(* IEC 61131-3 sources: POMIRTS_lab3/AS/Library/brsystem, 2 files *)

(* ---- brsystem.fun ---- *)
(********************************************************************
 * COPYRIGHT -- Bernecker + Rainer
 ********************************************************************
 * Library: brsystem
 * File: brsystem.fun
 * Author: B+R
 ********************************************************************
 * Functions and function blocks of library brsystem
 ********************************************************************)

FUNCTION_BLOCK MEMInfo				(*returns information about the memory areas available on the system*)
	VAR_INPUT
		enable	:BOOL;				(*enables execution*)
	END_VAR
	VAR_OUTPUT
		status	:UINT;				(*execution status: ERR_OK, ERR_FUB_ENABLE_FALSE, 0xXXXX = see help*)
		FreeUSR_Ram	:UDINT;			(*SG3: free memory in USER RAM SG4: free memory in SRAM (Userram)*)
		FreeSYSTEM	:UDINT;			(*SG3: free system memory SG4: not used, always 0*)
		FreeUSR_Prom	:UDINT;		(*SG3: free memory in USER PROM SG4: free memory of HD where RPSHD is located*)
		FreeSYS_Prom	:UDINT;		(*SG3: free memory in system PROM SG4: free memory of HD where RPSHD is located*)
		FreeFIX_Ram	:UDINT;			(*SG3: free memory in FIX RAM SG4: not used, always 0*)
		FreeTMP_Ram	:UDINT;			(*SG3: free temporary memory in RAM SG4: free memory in DRAM*)
		FreeMEMCARD	:UDINT;			(*SG3: free memory on MEMCARD SG4: not used, always 0*)
	END_VAR
END_FUNCTION_BLOCK

FUNCTION_BLOCK MEMxInfo				(*returns information about the memory areas available in the system; asynchronous execution*)
	VAR_INPUT
		enable	:BOOL;   			(*enables execution*)
		mem_typ	:UDINT;				(*memory type: brDRAM, brUSRRAM, brSYSROM, brUSRROM*)
	END_VAR
	VAR_OUTPUT
		status	:UINT;				(*execution status: ERR_OK, ERR_FUB_ENABLE_FALSE, ERR_FUB_BUSY, 0xXXXX = see help*)
		MemSize	:UDINT;				(*total memory size in bytes*)
		FreeMemSize	:UDINT;			(*size of available memory in bytes*)
		BiggestFreeBlockSize	:UDINT;	(*size of the largest available block in memory in bytes*)
	END_VAR
	VAR
		i_state	:UINT;				(*internal variable*)
		i_result	:UINT;			(*internal variable*)
		i_tmp	:UDINT;				(*internal variable*)
	END_VAR
END_FUNCTION_BLOCK

FUNCTION_BLOCK SysInfo				(*returns information about the target system*)
	VAR_INPUT
		enable	:BOOL;				(*enables execution*)
	END_VAR
	VAR_OUTPUT
		init_reason	:USINT;			(*reason for initialization*)
		init_count	:USINT;			(*SG3: the value is increased by every INIT (warm restart) SG4: not used, always 0*)
		tick_count	:UDINT;			(*tick count*)
		version	:UDINT;				(*operating system version of the target system*)
	END_VAR
END_FUNCTION_BLOCK

FUNCTION_BLOCK RTInfo				(*returns runtime information about the software object*)
	VAR_INPUT
		enable	:BOOL;				(*enables execution*)
	END_VAR
	VAR_OUTPUT
		status	:UINT;				(*execution status: ERR_OK, ERR_FUB_ENABLE_FALSE, 0xXXXX = see help*)
		cycle_time	:UDINT;			(*cycle time in microsec*)
		init_reason	:SINT;			(*reason for initialization*)
		task_class	:SINT;			(*task class (SG3: #1 - #4 SG4: #1 - #8)*)
	END_VAR
END_FUNCTION_BLOCK

FUNCTION_BLOCK TARGETInfo			(*returns information about the target system used*)
	VAR_INPUT
		enable	:BOOL;				(*enables execution*)
		pOSVersion	:UDINT;			(*string given as a pointer (min. 7 char), where the os version is written*)
	END_VAR
	VAR_OUTPUT
		status	:UINT;				(*execution status: ERR_OK, ERR_FUB_ENABLE_FALSE, 0xXXXX = see help*)
		DataFormat	:USINT;			(*wether "big endian" or "little endian" ("TARGET_BIG_ENDIAN"/"TARGET_LITTLE_ENDIAN")*)
	END_VAR
END_FUNCTION_BLOCK

FUNCTION_BLOCK HWInfo				(*returns information about the hardware configuration*)
	VAR_INPUT
		enable	:BOOL;				(*enables execution*)
		first	:BOOL;				(*determines the hardware module on which the FUB is used 0/1 next/first*)
		pName	:UDINT;				(*string given as a pointer, where the name of the module is written*)
	END_VAR
	VAR_OUTPUT
		status	:UINT;				(*execution status: ERR_OK, ERR_FUB_ENABLE_FALSE, 0xXXXX = see help*)
		family	:USINT;				(*family designation*)
		usetype	:USINT;				(*hardware type*)
		module_typ	:UDINT;			(*module type*)
		master_no	:USINT;			(*logical number of the IO master, RIO master, CAN bus with CANIO*)
		slave_no	:USINT;			(*slave number*)
		module_adr	:USINT;			(*hardware module address (decimal)*)
		slot_no	:USINT;				(*slot of the first submodule found (decimal)*)
	END_VAR
	VAR
		next_vw_p	:UDINT;			(*internal variable*)
		last_modul_p	:UDINT;		(*internal variable*)
		next_entry_p	:UDINT;		(*internal variable*)
		next_entry_ix	:USINT;		(*internal variable*)
		next_slot_ix	:USINT;		(*internal variable*)
		last_rio_master	:USINT;		(*internal variable*)
	END_VAR
END_FUNCTION_BLOCK

FUNCTION_BLOCK SysconfInfo			(*returns the parameters for a sysconf entry*)
	VAR_INPUT
		enable	:BOOL;				(*enables execution*)
		pEntry	:UDINT;				(*string given as a pointer, where the name of the entry is written*)
		pValue	:UDINT;				(*string given as a pointer, where the value of the entry is copied*)
		value_len	:UDINT;			(*length of the "value-string"*)
	END_VAR
	VAR_OUTPUT
		status	:UINT;				(*execution status: ERR_OK, ERR_FUB_ENABLE_FALSE, 0xXXXX = see help*)
	END_VAR
END_FUNCTION_BLOCK

FUNCTION_BLOCK SysconfSet			(*sets the parameters for a sysconf entry*)
	VAR_INPUT
		enable	:BOOL;				(*enables execution*)
		pEntry	:UDINT;				(*string given as a pointer, where the name of the entry is written*)
		pNewValue	:UDINT;			(*string given as a pointer, where the new value of the entry is written*)
		option	:USINT;				(*sets the parameter volatile/permanent ("brSYSCONF_SET_VOLATILE"/"brSYSCONF_SET_NON_VOLATILE")*)
	END_VAR
	VAR_OUTPUT
		status	:UINT;				(*execution status: ERR_OK, ERR_FUB_ENABLE_FALSE, 0xXXXX = see help*)
	END_VAR
END_FUNCTION_BLOCK

FUNCTION_BLOCK BatteryInfo			(*returns the state of the battery*)
	VAR_INPUT
		enable	:BOOL;				(*enables execution*)
		pDevice	:UDINT;				(*device name given as a pointer*)
	END_VAR
	VAR_OUTPUT
		status	:UINT;				(*execution status: ERR_OK, ERR_FUB_ENABLE_FALSE, 0xXXXX = see help*)
		state	:USINT;				(*state of the battery*)
	END_VAR
END_FUNCTION_BLOCK

FUNCTION_BLOCK EXCInfo				(*returns information about the software object that triggered the exception*)
	VAR_INPUT
		enable	:BOOL;				(*enables execution*)
	END_VAR
	VAR_OUTPUT
		status	:UINT;				(*execution status: ERR_OK, ERR_FUB_ENABLE_FALSE, 0xXXXX = see help*)
		task_class	:UDINT;			(*task class in which the exception was triggered*)
		task_ident	:UDINT;			(*ID number of the software object that triggered the exception*)
	END_VAR
END_FUNCTION_BLOCK

FUNCTION_BLOCK ZYKVLenable			(*enables/disables the cycle time monitoring of software objects*)
	VAR_INPUT
		enable	:BOOL;				(*enables execution*)
		mode	:BOOL;				(*0/1 monitoring off/on*)
	END_VAR
	VAR_OUTPUT
		status	:UINT;				(*execution status: ERR_OK, ERR_FUB_ENABLE_FALSE, 0xXXXX = see help*)
	END_VAR
END_FUNCTION_BLOCK

FUNCTION_BLOCK PMemGet				(*reads data of len byte from the permanent memeory area beginning at offset*)
	VAR_INPUT
		enable	:BOOL;				(*enables execution*)
		offset	:UDINT;				(*offset within the permanent memory area*)
		len	 :UDINT;				(*length of data area to be read*)
		adress	:UDINT;				(*address where the read data is copied*)
	END_VAR
	VAR_OUTPUT
		status	:UINT;				(*execution status: ERR_OK, ERR_FUB_ENABLE_FALSE, 0xXXXX = see help*)
	END_VAR
END_FUNCTION_BLOCK

FUNCTION_BLOCK PMemPut				(*writes len bytes to the permanent memory area beginning at offset*)
	VAR_INPUT
		enable	:BOOL;				(*enables execution*)
		offset	:UDINT;				(*offset within the permanent memory area*)
		len	 :UDINT;				(*length of data area to be written*)
		adress	:UDINT;				(*address of the data to be written to the permanent memory area*)
	END_VAR
	VAR_OUTPUT
		status	:UINT;				(*execution status: ERR_OK, ERR_FUB_ENABLE_FALSE, 0xXXXX = see help*)
	END_VAR
END_FUNCTION_BLOCK

FUNCTION_BLOCK PMemSize				(*determines the size of permanent memory area in its existing configuration*)
	VAR_INPUT
		enable	:BOOL;				(*enables execution*)
	END_VAR
	VAR_OUTPUT
		status	:UINT;				(*execution status: ERR_OK, ERR_FUB_ENABLE_FALSE, 0xXXXX = see help*)
		size	:UDINT;				(*size of permanent memory area*)
	END_VAR
END_FUNCTION_BLOCK

(* ---- brsystem.var ---- *)
(********************************************************************
 * COPYRIGHT -- Bernecker + Rainer
 ********************************************************************
 * Library: brsystem
 * File: brsystem.var
 * Author: B+R
 ********************************************************************
 * Local variables of library brsystem
 ********************************************************************)

VAR CONSTANT
	brSYSCONF_SET_NON_VOLATILE	: BOOL	:= TRUE;	(*set permanent value*)
	brERR_INVALID_PARAMETER	: UINT	:= 27251;		(*invalid parameter transferred*)
	brSYSCONF_SET_VOLATILE	: BOOL	:= FALSE;		(*set non-permanent value*)
	INIT_REASON_WARMSTART	: SINT	:= 1;			(*warm restart boot information*)
	INIT_REASON_COLDSTART	: SINT	:= 2;			(*cold restart boot information*)
	brERR_INVALID_DEVICE	: UINT	:= 27250;		(*battery monitoring*)
	brAUTOMATION_RUNTIME	: USINT	:= 4;			(*series recognition*)
	TARGET_LITTLE_ENDIAN	: USINT	:= 1;			(*formatSpec*)
	INIT_REASON_DOWNLOAD	: SINT	:= 3;			(*download boot information*)
	INIT_REASON_UNKNOWN	: SINT	:= -1;				(*unknown boot information*)
	brBATTERY_MISSING	: USINT	:= 3;				(*battery monitoring*)
	TARGET_BIG_ENDIAN	: USINT	:= 2;				(*formatSpec*)
	brBATTERY_NOTEST	: USINT	:= 2;				(*battery monitoring*)
	brSYSTEM_MODULE	: USINT	:= 2;					(*usage recognition*)
	brPLUGIN_MODULE	: USINT	:= 10;					(*usage recognition*)
	brLOGICSCANNER	: USINT	:= 3;					(*series recognition*)
	brBATTERY_LOW	: USINT	:= 0;					(*battery monitoring*)
	brPOWERPANEL	: USINT	:= 5;					(*series recognition*)
	brBATTERY_OK	: USINT	:= 1;					(*battery monitoring*)
	brREMOTE_IO	: USINT	:= 4;						(*usage recognition*)
	brNO_FAMILY	: USINT	:= 255;						(*series recognition*)
	brETHER_IO	: USINT	:= 6;						(*usage recognition*)
	brPRODUCT	: USINT	:= 0;						(*usage recognition*)
	brBASE_IO	: USINT	:= 3;						(*usage recognition*)
	brCAN_IO	: USINT	:= 5;						(*usage recognition*)
	brACOPOS	: USINT	:= 7;						(*usage recognition*)
	brUSRRAM	: UDINT	:= 1;						(*USRRAM memory type*)
	brSYSROM	: UDINT	:= 2;						(*SYSROM memory type*)
	brUSRROM	: UDINT	:= 3;						(*USRROM memory type*)
	brLOCAL_REMANENT_PV  : UDINT	:= 4;			(*local REMMEM memory type*)
	brGLOBAL_REMANENT_PV : UDINT	:= 5;			(*global REMMEM memory type*)
	brPANEL	: USINT	:= 6;							(*series recognition*)
	brADDON	: USINT	:= 7;							(*series recognition*)
	brC300	: USINT	:= 8;							(*series recognition*)
	brC200	: USINT	:= 9;							(*series recognition*)
	br2010	: USINT	:= 0;							(*series recognition*)
	br2005	: USINT	:= 1;							(*series recognition*)
	br2003	: USINT	:= 2;							(*series recognition*)
	brDRAM	: UDINT	:= 0;							(*DRAM memory type*)
	brKEY	: USINT	:= 8;							(*usage recognition*)
	brCPU	: USINT	:= 1;							(*usage recognition*)
	brPP	: USINT	:= 255;							(*usage recognition*)
	brX2X	: USINT	:= 10;							(*series recognition*)
END_VAR
